Fanuc KAREL source: KT00929.KL

PROGRAM KT00929
%NOLOCKGROUP
VAR
  I1: INTEGER
  I2: INTEGER
  OUT: INTEGER
BEGIN
  I1 = 2
  I2 = 3
  I1 = 2
  I2 = 3
  OUT = ORD(I1, 1)
END KT00929
